TYPE "FRK_TestStatus"
VERSION : 0.1
   STRUCT
      "Done" : Bool;
      "Checks" : Int;
      "Failures" : Int;
      "FirstFailure" : Int;
      "ImageHash" : Array[0..7] of DWord;
   END_STRUCT;
END_TYPE
